Fanuc KAREL source: kc00034.KL

-- PROVISIONAL review KL for V770-1; original PC SHA256 afee188c7fd105cb94df7323e4570702abd040e3b405629d0c3952ba107a0f34
-- Incomplete behavior may be omitted. Consult companion uncertainty JSON. Do not deploy.
PROGRAM KC00034
%NOLOCKGROUP
BEGIN
  -- UNRESOLVED_PC offsets 5-29; opcodes 27,22,22,2A,22,31
  -- UNRESOLVED_PC offsets 34-38; opcodes 7F
END KC00034
